FUNCTION_BLOCK PUBLIC FB_Filling EXTENDS FB_SFC_Cycle IMPLEMENTS ITF_FB_SFC_Cycle
VAR_INPUT
	valFilling				: E_Pis_Name	;
	setWeight				: REAL:=200.0;	//kg
	actWeight				: REAL:=100.0;	//kg
	Tolerance				: REAL:=0.5;	//kg
	
END_VAR
VAR
	fbPis					: FB_Piston;	
	stPis_Filling			: REFERENCE TO ST_Piston;
	
	MinWeight	: REAL;
	MaxWeight	: REAL;
	
	reqTara		: BOOL;

END_VAR
VAR_IN_OUT
	eFill_State				: E_Filling_State;
END_VAR
VAR_OUTPUT
	eFill_State_HMI			: E_Filling_State;
	pumpFilling				: BOOL;
END_VAR

act_GetReference();

act_Oper();

MinWeight:=setWeight-Tolerance;
MaxWeight:=setWeight+Tolerance;
eFill_State_HMI:=eFill_State;

IF reqTara THEN;
	IF m_Tara() THEN;
		reqTara:=FALSE;
	ELSE;
		// tara command in process
	END_IF
END_IF

ACTION _aCheck_Condition_active:
// communication to weight


// check tara == weghit value <= 0.5 kg and >= -0.5 kg ==> 0 +- 0.5
bStepDone:=FALSE;
IF TRUE
//AND actWeight >= -0.5 AND actWeight <= 0.5 
AND actWeight < MinWeight 
AND eFill_State=E_Filling_State.eReady_ToFill
AND TRUE
THEN;
	bStepDone:=TRUE;
END_IF
END_ACTION

ACTION _aFilling_Process_active:
// check frow weight >= min value from recipe

pumpFilling:=m_FillingActive(); // Run autofiling process...
eFill_State:=E_Filling_State.eFilling_InProcess;

bStepDone:=FALSE;
IF actWeight >= MinWeight THEN;
	bStepDone:=TRUE;
END_IF
END_ACTION

ACTION _aFilling_Process_entry:
// open filling valve
fbPis.m_SetByRecipe(stPis:=stPis_Filling, 			req:=E_Piston_Recipe_State.Act);
// run pump
END_ACTION

ACTION _aFilling_Process_exit:
// close valve

// stop pump
END_ACTION

ACTION _aNo_Condition_active:
// print error
END_ACTION

ACTION _aReset_entry:
//close filing valve 
fbPis.m_SetByRecipe(stPis:=stPis_Filling, 			req:=E_Piston_Recipe_State.Release);

pumpFilling:=FALSE;
IF eFill_State=E_Filling_State.eFilling_InProcess THEN;
	eFill_State:=E_Filling_State.eReady_ToFill;
END_IF
bRun:=FALSE;
END_ACTION

ACTION act_GetReference:
m_Set_SFCFlags_Reference();

stPis_Filling				REF= g_Piston.stPis[valFilling];

(*
stPis_TankB				REF= g_Piston.stPis[valTankB];
stPis_TapWater			REF= g_Piston.stPis[valTapWater];
stPis_TapWater_else		REF= g_Piston.stPis[valTapWater_else];
stPis_TapWater_Drain	REF= g_Piston.stPis[valTapWater_Drain];
stPis_BlockWater		REF= g_Piston.stPis[valBlockWater];
stPis_WaterSource		REF= g_Piston.stPis[valWaterSource];
stPis_WaterSource_Drain	REF= g_Piston.stPis[valWaterSource_Drain];
stPis_Drain				REF= g_Piston.stPis[valDrain];
stPis_CIP				REF= g_Piston.stPis[valCIP];
stPis_CIP_Sel			REF= g_Piston.stPis[valCIP_Sel];
*)
END_ACTION

ACTION act_Oper:
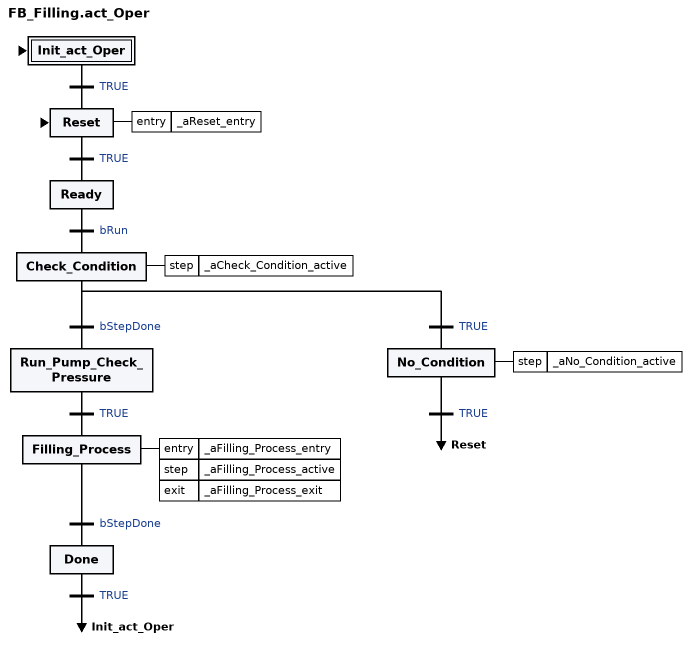
INITIAL_STEP Init_act_Oper:
END_STEP
TRANSITION FROM Init_act_Oper TO Reset
    := TRUE;
END_TRANSITION
STEP Reset:
    _aReset_entry(P1);  // entry action
END_STEP
TRANSITION FROM Reset TO Ready
    := TRUE;
END_TRANSITION
STEP Ready:
END_STEP
TRANSITION FROM Ready TO Check_Condition
    := bRun;
END_TRANSITION
STEP Check_Condition:
    _aCheck_Condition_active(N);  // step action
END_STEP
TRANSITION FROM Check_Condition TO Run_Pump_Check_Pressure
    := bStepDone;
END_TRANSITION
STEP Run_Pump_Check_Pressure:
END_STEP
TRANSITION FROM Run_Pump_Check_Pressure TO Filling_Process
    := TRUE;
END_TRANSITION
STEP Filling_Process:
    _aFilling_Process_entry(P1);  // entry action
    _aFilling_Process_active(N);  // step action
    _aFilling_Process_exit(P0);  // exit action
END_STEP
TRANSITION FROM Filling_Process TO Done
    := bStepDone;
END_TRANSITION
STEP Done:
END_STEP
TRANSITION FROM Done TO Init_act_Oper
    := TRUE;
END_TRANSITION
TRANSITION FROM Check_Condition TO No_Condition
    := TRUE;
END_TRANSITION
STEP No_Condition:  // min time T#2s
    _aNo_Condition_active(N);  // step action
END_STEP
TRANSITION FROM No_Condition TO Reset
    := TRUE;
END_TRANSITION
// branch label Branch0_act_Oper
END_ACTION

METHOD m_FillingActive : BOOL
VAR_INPUT
END_VAR

actWeight:=actWeight+0.1;
m_FillingActive:=TRUE;
END_METHOD

{warning 'add method implementation '}
METHOD m_Set_SFCFlags_Reference : BOOL
//Set reference to SFC flags

refSFC.SFCInit REF= SFCInit;
refSFC.SFCReset REF= SFCReset;
refSFC.SFCError REF= SFCError;
refSFC.SFCEnableLimit REF= SFCEnableLimit;
refSFC.SFCErrorStep REF= SFCErrorStep;
refSFC.SFCErrorPOU REF= SFCErrorPOU;
refSFC.SFCQuitError REF= SFCQuitError;
refSFC.SFCPause REF= SFCPause;
refSFC.SFCTrans REF= SFCTrans;
refSFC.SFCCurrentStep REF= SFCCurrentStep;
refSFC.SFCTip REF= SFCTip;
refSFC.SFCTipMode REF= SFCTipMode;

// Cycle handle for SFC
m_SFC_Handle();
END_METHOD

METHOD m_Tara : BOOL
VAR_INPUT
END_VAR
actWeight:=0.0;
m_Tara:=TRUE;
END_METHOD

END_FUNCTION_BLOCK

(* stored: Version 1.1.0.1, ProductVersion 3.1.4024.15
   POU FB_Filling: Id {57ce42fe-7c67-4e80-b858-2c5ec698a104}, SpecialFunc None
   Action _aCheck_Condition_active: Id {52e30844-68a2-4937-9c55-054be0048d36}
   Action _aFilling_Process_active: Id {86a344ec-4f3b-47c2-bf07-c3fd927019f9}
   Action _aFilling_Process_entry: Id {a4bdcf2a-7b2e-4685-bd70-7299b1106ef5}
   Action _aFilling_Process_exit: Id {a37338e0-afaf-4228-9a18-d54bc1b114a9}
   Action _aNo_Condition_active: Id {f128ce1d-c88a-4f8d-8acc-62baade13eee}
   Action _aReset_entry: Id {11253cd7-8b45-408b-91df-74590fbcd973}
   Action act_GetReference: Id {cd6f94bf-aa3a-47a2-b52c-08d8cae50358}
   Action act_Oper: Id {9cd67642-f4cb-42e4-9826-dae8e9f291a1}
   Method m_FillingActive: Id {e50ac11a-8566-4bd3-8e9e-4ca51d09cfb6}
   Method m_Set_SFCFlags_Reference: Id {72f7dfaa-0d20-44b1-86c3-1f73dee8a36f}
   Method m_Tara: Id {d585ec45-9719-4ad3-b51d-9430cbc3ebd5} *)
